(* Production-style program with a FB_LIC nested in FB_LICInitHost. It follows
   PRG_ATMInit: one motor, the PMPS state-name configurators and the host. The
   arbiter, fast-fault output, persistent storage and DB reader are shared in
   GVL_PRG and ticked by PRG_PMPS_PRE and PRG_PMPS_POST. The configurators are in
   the PRG, because the host's references are not bound yet when its
   declaration initialisers run. The PMPS DB is plc-cc-motion.json. *)
PROGRAM PRG_LIC
VAR
    {attribute 'TcNcAxis' := 'PRG_LIC_Y'}
    axRef         : AXIS_REF;
    fbMotor       : FB_MotionStageNC(
        AxisRef                := axRef,
        iPersistentDataStorage := GVL_PRG.fbPDS,
        sName                  := 'LICINIT'
    );
    aiMotionStage : ARRAY[1..MotionConstants.MAX_STATE_MOTORS] OF I_MotionStage := [fbMotor];

    astPositionState : ARRAY[1..MotionConstants.MAX_STATE_MOTORS]
                         OF ARRAY[1..GeneralConstants.MAX_STATES] OF ST_PositionState;
    stDefault : ST_PositionState := (
        bMoveOk       := TRUE,
        bValid        := TRUE,
        bUseRawCounts := FALSE
    );
    afbStatePMPS : ARRAY[1..4] OF FB_CC_StatePMPSConfig[
        (stPositionState := astPositionState[1][E_LIC_States.OUT],
         stDefault       := stDefault,
         fPosition       := 10,
         sPmpsState      := 'TST:LIC-OUT'),
        (stPositionState := astPositionState[1][E_LIC_States.MIRROR1],
         stDefault       := stDefault,
         fPosition       := 20,
         sPmpsState      := 'TST:LIC-MIRROR1'),
        (stPositionState := astPositionState[1][E_LIC_States.MIRROR2],
         stDefault       := stDefault,
         fPosition       := 30,
         sPmpsState      := 'TST:LIC-MIRROR2'),
        (stPositionState := astPositionState[1][E_LIC_States.TARGET],
         stDefault       := stDefault,
         fPosition       := 40,
         sPmpsState      := 'TST:LIC-TARGET')
    ];

    fbHost : FB_LICHost(
        aiMotionStage         := aiMotionStage,
        astPositionState      := astPositionState,
        fbFFHWO               := GVL_PRG.fbFastFaultOutput1,
        fbArbiter             := GVL_PRG.fbArbiter1,
        sDeviceName           := 'TST:LIC',
        sTransitionKey        := 'TST:LIC-TRANSITION',
        bEnableBeamParams     := TRUE,
        bEnablePositionLimits := TRUE,
        bReadDBNow            := TRUE,
        bFileReaderBusy       := MOTION_GVL.fbPmpsFileReader.bBusy,
        bFileReaderError      := MOTION_GVL.fbPmpsFileReader.bError
    );

    i          : UINT;
    bFirstScan : BOOL := TRUE;
END_VAR

IF bFirstScan THEN
    fbMotor.SetModeEnableLimits(
        LimBackward    := TRUE,
        LimForward     := TRUE,
        HomeEnable     := FALSE,
        BrakeMode      := E_StageBrakeMode.IF_ENABLED,
        EnableMode     := E_StageEnableMode.DURING_MOTION,
        HomeMode       := E_EpicsHomeCmd.LOW_LIMIT,
        UserEnable     := TRUE,
        HardwareEnable := TRUE
    );
    fbMotor.SetVelocity(
        Velocity := 15.5
    );
    fbMotor.RestoreMotionParams      := FALSE;
    fbMotor.DoNotRestoreNcParameters := TRUE;
    bFirstScan := FALSE;
END_IF

FOR i := 1 TO 4 DO
    afbStatePMPS[i]();
END_FOR

fbHost();
fbMotor();

END_PROGRAM

(* stored: Version 1.1.0.1
   POU PRG_LIC: Id {87bd08e1-1b74-4d3f-9958-0766e50a089d}, SpecialFunc None *)
